(* IEC 61131-3 sources: plcassist-cli/packages/volt-lsp-iec/test-corpus/awa-palletizer/Device/Plc Logic/Application/Library Manager/(unresolved)/cmpusermgr interfaces, 4 files *)

(* ---- AUDITINFOIDS.gvl ---- *)
VAR_GLOBAL
	AUDIT_INFOID_USER_LOCKED : DINT := 16#1;
END_VAR

(* ---- CONSTANTS.gvl ---- *)
VAR_GLOBAL
	USERMGR_RIGHT_NONE : DWORD := 0;
	USERMGR_RIGHT_VIEW : DWORD := 1;
	USERMGR_RIGHT_MODIFY : DWORD := 2;
	USERMGR_RIGHT_EXECUTE : DWORD := 4;
	USERMGR_RIGHT_ADD_REMOVE : DWORD := 8;
	USERMGR_RIGHT_OEM : DWORD := 16#FF000000;
	USERMGR_RIGHT_ALL : DWORD := 16#FFFFFFFF;
END_VAR

(* ---- EVENTIDS.gvl ---- *)
VAR_GLOBAL
	CMPID_CMPUSERMGR : DWORD := 16#61;
	EVTPARAMID_CMPUSERMGRDATABASECHANGED : WORD := 16#1;
	EVTVERSION_CMPUSERMGRDATABASECHANGED : WORD := 16#1;
	EVT_USERMGRDATABASECHANGED : DWORD := (SHL(UINT_TO_DWORD(EVTCLASS_INFO), 16) OR 16#1);
	EVTPARAMID_CMPUSERMGRPASSWORDVALIDITY : WORD := 16#3;
	EVTVERSION_CMPUSERMGRPASSWORDVALIDITY : WORD := 16#1;
	EVT_USERMGRPASSWORDVALIDITY : DWORD := (SHL(UINT_TO_DWORD(EVTCLASS_INFO), 16) OR 16#5);
	EVT_USERMGRPASSWORDEXPIRED : DWORD := (SHL(UINT_TO_DWORD(EVTCLASS_WARNING), 16) OR 16#6);
END_VAR

(* ---- PROPERTIES.gvl ---- *)
VAR_GLOBAL
	USERMGR_USER_PROP_PASSWORD_EXPIRED : DWORD := 16#1000;
	USERMGR_USER_PROP_ALLOW_CHANGE_PASSWORD : DWORD := 16#2000;
	USERMGR_USER_PROP_DEFAULT : DWORD := (USERMGR_USER_PROP_ALLOW_CHANGE_PASSWORD + USERMGR_USER_PROP_PASSWORD_EXPIRED);
END_VAR
